// TIA Portal V19 export
// export: Created 2026-10-15T09:44:23.177447Z, ExportSetting WithDefaults, DisplayName Totally Integrated Automation Portal, DisplayVersion V19, DisplayName TIA Portal Openness, DisplayVersion V19, DisplayName TIA Portal Version Control Interface, DisplayVersion V19, DisplayName STEP 7 Professional, DisplayVersion V19, DisplayName STEP 7 Safety, DisplayVersion V19, DisplayName WinCC Basic/Comfort/Advanced, DisplayVersion V19, DisplayName WinCC Unified, DisplayVersion V19
FUNCTION "ROLL_AdvanceTime" : Void   // FC9, SCL
{ S7_Optimized_Access := 'TRUE' }
VERSION : 0.1
// stored: AutoNumber true, IsIECCheckEnabled false, SetENOAutomatically false, UDAEnableTagReadback false
   VAR_INPUT
      DeltaMs : LReal;
   END_VAR
   VAR_TEMP
      n : Int;
   END_VAR
BEGIN

   IF #DeltaMs < 0.0 THEN
       "ROLL_IO".ConversionFault := TRUE;
       RETURN;
   END_IF;
   FOR #n := 0 TO 127 DO
       IF "ROLL_State".S5Timers[#n].RemainingMs > 0.0 THEN
           "ROLL_State".S5Timers[#n].RemainingMs := "ROLL_State".S5Timers[#n].RemainingMs - #DeltaMs;
           IF "ROLL_State".S5Timers[#n].RemainingMs <= 0.0 THEN
               "ROLL_State".S5Timers[#n].RemainingMs := 0.0;
               "ROLL_State".S5Timers[#n].Q := "ROLL_State".S5Timers[#n].Mode = 0;
           END_IF;
       END_IF;
   END_FOR;
   "ROLL_IO".ClockMs := "ROLL_IO".ClockMs + #DeltaMs;
   WHILE "ROLL_IO".ClockMs >= 250.0 DO
       "ROLL_IO".ClockMs := "ROLL_IO".ClockMs - 250.0;
       "ROLL_State".M[3, 4] := NOT "ROLL_State".M[3, 4];
       IF NOT "ROLL_State".M[3, 4] THEN
           "ROLL_State".M[3, 5] := NOT "ROLL_State".M[3, 5];
           IF NOT "ROLL_State".M[3, 5] THEN
               "ROLL_State".M[3, 6] := NOT "ROLL_State".M[3, 6];
               IF NOT "ROLL_State".M[3, 6] THEN
                   "ROLL_State".M[3, 7] := NOT "ROLL_State".M[3, 7];
               END_IF;
           END_IF;
       END_IF;
   END_WHILE;
END_FUNCTION
